(*
SPDX-License-Identifier: MIT
License: https://opensource.org/license/mit
*)

(*!
<summary>Owns the pending multi-cycle test used for deadline verification.</summary>
<description>
Owns persistent child storage and fixed parent associations. Use in one task without reentry.
Children is borrowed and must not be modified by application code. Constructor callbacks are not used.
</description>
*)

{attribute 'no_assign'}
{attribute 'no_explicit_call' := 'do not call this function block directly'}
FUNCTION_BLOCK DeadlineTestGroup EXTENDS TOF_Testing.TestGroup<1>
VAR_STAT
	//! <summary>Class name shared by all instances of this function block.</summary>
	{attribute 'hide'}
	_ClassName : STRING := __POUNAME();
END_VAR
VAR
	{attribute 'hide'}
	{attribute 'init_namespace'}
	_NamespaceName : STRING;
END_VAR
VAR_OUTPUT
	//! <summary>Owned multi-cycle leaf with an externally selected deadline.</summary>
	Child : AssertionIsolationProbe(name := "Deadline", parent := THIS^);
END_VAR
VAR
	_Children : ARRAY [0.._ChildCount - 1] OF TOF_Testing.ITestElement :=
	[
		Child
	];
END_VAR

//! <summary>Borrows the concrete class name for the lifetime of this instance; callers must not modify it.</summary>
{attribute 'monitoring' := 'call'}
PROPERTY ClassName : REFERENCE TO STRING
GET
ClassName REF= _ClassName;
END_GET
END_PROPERTY

//! <summary>Borrows the compiler-initialized namespace; callers must not modify the returned reference.</summary>
{attribute 'monitoring' := 'call'}
PROPERTY NamespaceName : REFERENCE TO STRING
GET
NamespaceName REF= _NamespaceName;
END_GET
END_PROPERTY

//! <summary>Reports the complete concrete instance size, excluding separately allocated storage.</summary>
{attribute 'monitoring' := 'call'}
PROPERTY SelfSize : ULINT
GET
SelfSize := XSIZEOF(THIS^);
END_GET
END_PROPERTY

//! <summary>Borrows the fixed array of this concrete group; do not modify it.</summary>
{attribute 'monitoring' := 'call'}
PROPERTY Children : REFERENCE TO ARRAY [0.._ChildCount - 1] OF TOF_Testing.ITestElement
GET
Children REF= _Children;
END_GET
END_PROPERTY

END_FUNCTION_BLOCK

(* stored: Version 1.1.0.1
   POU DeadlineTestGroup: Id {6c4452db-0c67-4997-acb6-51697d5a2829}, SpecialFunc None
   Property ClassName: Id {8999a2aa-2eee-4317-9814-7943d215ade1}
   Get Get: Id {e8b09d0d-078d-4cfa-91b5-5411d475116f}
   Property NamespaceName: Id {2f284129-2402-46a5-b874-d38f3f6bc0c3}
   Get Get: Id {fc9261b0-9ca9-40bb-b13b-86390a707f49}
   Property SelfSize: Id {ad5e4443-1eba-49ab-9931-83053b31010d}
   Get Get: Id {65a239a0-0440-4a65-86f1-25933594997d}
   Property Children: Id {4084a0e6-a024-4d89-b82e-5449c4ed942e}
   Get Get: Id {f4a34b41-ce67-45b7-bd17-0988cf40b3db} *)
